PROGRAM main
  VAR
    SA1 AT %IX0.0 : BOOL; (* mano izquierda *)
    SA2 AT %IX0.1 : BOOL; (* mano derecha *)
    SA3 AT %IX0.2 : BOOL; (* tercera mano *)
    H1 AT %QX0.0  : BOOL; (* prensa *)
    H2 AT %QX0.1  : BOOL;
    H3 AT %QX0.2  : BOOL;
    H5 AT %QX0.4  : BOOL;
  END_VAR
  VAR  (* added by the conversion: wires and edge detectors of the diagram *)
    _AND1_OUT : BOOL;
    _OR6_OUT : BOOL;
    _NOT10_OUT : BOOL;
    _NOT15_OUT : BOOL;
    _AND13_OUT : BOOL;
  END_VAR

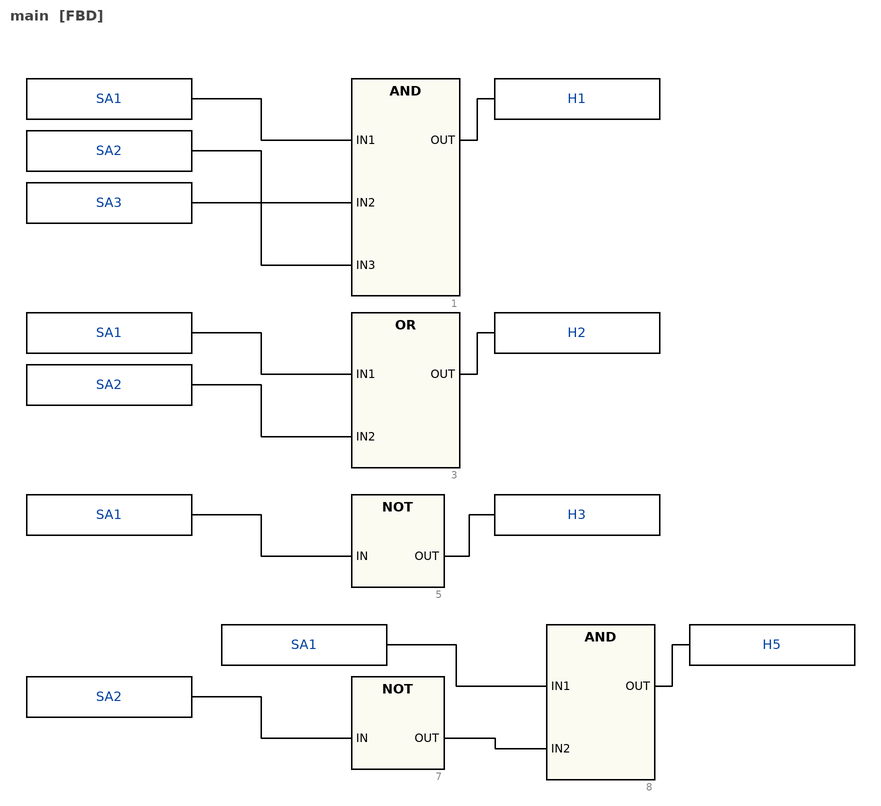
(* FBD diagram, written out as Structured Text *)
_AND1_OUT := SA1 AND SA2 AND SA3;
H1 := _AND1_OUT;
_OR6_OUT := SA1 OR SA2;
H2 := _OR6_OUT;
_NOT10_OUT := NOT SA1;
H3 := _NOT10_OUT;
_NOT15_OUT := NOT SA2;
_AND13_OUT := SA1 AND _NOT15_OUT;
H5 := _AND13_OUT;
END_PROGRAM
